{region 'Documentation'}
(*!
<summary>Check that IN is strictly later than Minimum.</summary>
*)
{endregion}
FUNCTION_BLOCK AssertLaterThan_LDT EXTENDS AssertionBase
VAR_INPUT
    IN : LDT; //! Actual value checked or observed by this Assertion.
    Minimum : LDT; //! Exclusive lower bound; the actual value or count must be greater.
END_VAR

SUPER^();

{region 'Documentation'}
(*!
<summary>Evaluate the typed temporal relation and report higher-priority errors first.</summary>
*)
{endregion}
METHOD PROTECTED Assert
VAR
    Message : STRING(GVL_Constants.MessageLength);
    MinimumText : STRING(GVL_Constants.AssertionValueLength);
    ActualText : STRING(GVL_Constants.AssertionValueLength);
END_VAR
IF NOT EvaluationActive THEN
    RETURN;
END_IF;

IF Result = E_Result.Error THEN
    RETURN;
END_IF;

IF Result = E_Result.Failed THEN
    RETURN;
END_IF;

IF IN <= Minimum THEN
    MinimumText := LDT_TO_STRING(Minimum);
    ActualText := LDT_TO_STRING(IN);
    Message := CONCAT('Assertion failed: value is not later than limit. Minimum = ',
        MinimumText);
    Message := CONCAT(Message, ', Actual = ');
    Message := CONCAT(Message, ActualText);
    Message := CONCAT(Message, '.');
    Fail(Message := Message);
    RETURN;
END_IF;

Pass();
END_METHOD

END_FUNCTION_BLOCK

(* stored: Version 1.1.0.1
   POU AssertLaterThan_LDT: Id {0714e888-2406-4011-9de3-a62314ac4650}, SpecialFunc None
   Folder Internal: Id {57393b1b-028c-4de3-a0b2-5257b2c4c35a}
   Method Assert: Id {5772b5de-ae03-42c5-bb36-6fcfaf35907d} *)
